(* IEC 61131-3 sources: SRCI_CLIENT_PLC/RobotLibrary/Library/POUs/SuperImposing/MC_MoveSuperImposedDynamic/Structures, 4 files *)

(* ---- MoveSuperImposedDynamicOutCmd.st ---- *)
{attribute 'pack_mode' := '1'}
// -------------------------------------------------------------------------
//  SRCI Robot Library
// -------------------------------------------------------------------------
//
//  Object:      MoveSuperImposedDynamicOutCmd
//  Author:      Thorsten Brach
//  Date:        2024-08-01
//
//  Description:
//
//
//  Copyright:
//    (C) 2024 Thorsten Brach. All rights reserved
//             Licensed under the MIT License.
//
//  Disclaimer:
//    This project is provided without any guarantee and can be used for
//    private and commercial purposes. Any use is at the user’s
//    own risk and responsibility.
//
// -------------------------------------------------------------------------
TYPE MoveSuperImposedDynamicOutCmd :
STRUCT
  /// Distance-to-go [mm] of the current job
  /// • -1: No valid value because move command is not yet active (valid values are pending) or not supported by RC
  /// • >0: Actual distance between current and target position
  /// •  0: Target position reached
  RemainingDistance  : REAL;
  /// Percentage of already traversed superimposed offset.
  /// If not supported : • -1
  Progress           : REAL;
  /// TRUE if the offset for superimposed positioning is reached.
  OffsetReached      : BOOL;
END_STRUCT
END_TYPE

(* ---- MoveSuperImposedDynamicParCmd.st ---- *)
{attribute 'pack_mode' := '1'}
// -------------------------------------------------------------------------
//  SRCI Robot Library
// -------------------------------------------------------------------------
//
//  Object:      MoveSuperImposedDynamicParCmd
//  Author:      Thorsten Brach
//  Date:        2024-08-01
//
//  Description:
//
//
//  Copyright:
//    (C) 2024 Thorsten Brach. All rights reserved
//             Licensed under the MIT License.
//
//  Disclaimer:
//    This project is provided without any guarantee and can be used for
//    private and commercial purposes. Any use is at the user’s
//    own risk and responsibility.
//
// -------------------------------------------------------------------------
TYPE MoveSuperImposedDynamicParCmd :
STRUCT
  /// Additional distance and orientation for superimposed positioning
  Offset             : RobotCartesianPosition;
  /// Defines type of reference coordinate system of the offset position.
  ReferenceType      : ReferenceType;
  /// Value of the maximum velocity difference of the additional motion (not necessary reached).
  /// • > 0% Use specified value.
  /// • ≤ 0% Use the velocity defined by the move command that is superimposed. If no motion is active, use internal minimal velocity. (default)
 /// See chapter 5.5.7 Robot dynamics
  VelocityDiffRate   : REAL;
  /// Value of the maximum acceleration difference of the additional motion (not necessary reached).
  ///  •  <0% Use default acceleration (default)
  ///  •   0% Use internal minimal acceleration
  ///  • 100% Use maximal reference acceleration
  /// See chapter 5.5.7 Robot dynamics
  AccelerationDiffRate: REAL := -1.0; // ST-FIX F156: spec 6.3.30 / 6.3.31: '<0 %: use default (default)'
  /// Value of the maximum deceleration difference of the additional motion (not necessary reached).
  /// •  <0% Use default deceleration (default)
  /// •   0% Use internal minimal deceleration
  /// • 100% Use maximal reference deceleration
  /// See chapter 5.5.7 Robot dynamics
  DecelerationDiffRate: REAL := -1.0; // ST-FIX F156: spec 6.3.30 / 6.3.31: '<0 %: use default (default)'
  /// Value of the maximum jerk difference of the additional motion (not necessary reached).
  /// •  <0% Use default jerk (default)
  /// •   0% Use internal minimal jerk
  /// • 100% Use maximal reference jerk
  /// See chapter 5.5.7 Robot dynamics
  JerkDiffRate        : REAL := -1.0; // ST-FIX F156: spec 6.3.30 / 6.3.31: '<0 %: use default (default)'
  /// Index of tool
  /// •      0: Flange (default)
  /// • 1..254: Tool frames
  ToolNo             : USINT;
  /// Index of frame
  /// •      0: WCS (default)
  /// • 1..254: User frames
  FrameNo            : USINT;
  /// Define the interpolation mode for the superimposed motion
  InterpolationMode  : InterpolationMode;
END_STRUCT
END_TYPE

(* ---- MoveSuperImposedDynamicRecvData.st ---- *)
{attribute 'pack_mode' := '1'}
// -------------------------------------------------------------------------
//  SRCI Robot Library
// -------------------------------------------------------------------------
//
//  Object:      MoveSuperImposedDynamicRecvData
//  Author:      Thorsten Brach
//  Date:        2024-08-01
//
//  Description:
//
//
//  Copyright:
//    (C) 2024 Thorsten Brach. All rights reserved
//             Licensed under the MIT License.
//
//  Disclaimer:
//    This project is provided without any guarantee and can be used for
//    private and commercial purposes. Any use is at the user’s
//    own risk and responsibility.
//
// -------------------------------------------------------------------------
TYPE MoveSuperImposedDynamicRecvData EXTENDS RspHeader :
STRUCT
  /// Percentage of already traversed distance of current job.
  /// If not supported : • -1
  Progress          : UINT;
  /// Distance-to-go of the current job.
  /// • -1: No valid value because move command is not yet active (valid values are pending) or not supported by RC
  /// • >0: Actual distance between current and target position
  /// •  0: Target position reached
  RemainingDistance  : REAL;
  /// TRUE if the offset for superimposed positioning is reached.
  OffsetReached      : BOOL;
END_STRUCT
END_TYPE

(* ---- MoveSuperImposedDynamicSendData.st ---- *)
{attribute 'pack_mode' := '1'}
// -------------------------------------------------------------------------
//  SRCI Robot Library
// -------------------------------------------------------------------------
//
//  Object:      MoveSuperImposedDynamicSendData
//  Author:      Thorsten Brach
//  Date:        2024-08-01
//
//  Description:
//
//
//  Copyright:
//    (C) 2024 Thorsten Brach. All rights reserved
//             Licensed under the MIT License.
//
//  Disclaimer:
//    This project is provided without any guarantee and can be used for
//    private and commercial purposes. Any use is at the user’s
//    own risk and responsibility.
//
// -------------------------------------------------------------------------
TYPE MoveSuperImposedDynamicSendData EXTENDS CmdHeader:
STRUCT
  /// Value of the maximum velocity difference of the additional motion (not necessary reached).
  /// • > 0% Use specified value.
  /// • ≤ 0% Use the velocity defined by the move command that is superimposed. If no motion is active, use internal minimal velocity. (default)
 /// See chapter 5.5.7 Robot dynamics
  VelocityDiffRate    : UINT;
  /// Value of the maximum acceleration difference of the additional motion (not necessary reached).
  ///  •  <0% Use default acceleration (default)
  ///  •   0% Use internal minimal acceleration
  ///  • 100% Use maximal reference acceleration
  /// See chapter 5.5.7 Robot dynamics
  AccelerationDiffRate: UINT;
  /// Value of the maximum deceleration difference of the additional motion (not necessary reached).
  /// •  <0% Use default deceleration (default)
  /// •   0% Use internal minimal deceleration
  /// • 100% Use maximal reference deceleration
  /// See chapter 5.5.7 Robot dynamics
  DecelerationDiffRate: UINT;
  /// Value of the maximum jerk difference of the additional motion (not necessary reached).
  /// •  <0% Use default jerk (default)
  /// •   0% Use internal minimal jerk
  /// • 100% Use maximal reference jerk
  /// See chapter 5.5.7 Robot dynamics
  JerkDiffRate        : UINT;
  /// Index of tool
  /// •      0: Flange (default)
  /// • 1..254: Tool frames
  ToolNo              : USINT;
  /// Index of frame
  /// •      0: WCS (default)
  /// • 1..254: User frames
  FrameNo             : USINT;
  /// Reserve X
  Reserve_X           : REAL;
  /// Additional distance and orientation for superimposed positioning
  Offset              : RobotCartesianPosition;
  /// Defines type of reference coordinate system of the offset position.
  ReferenceType       : USINT;
  /// Define the interpolation mode for the superimposed motion
  InterpolationMode   : USINT;
END_STRUCT
END_TYPE
